FUNCTION_BLOCK STRING_TO_CAN_MSG (* STRING (bis 8 Zeichen) in eine CAN_MSG fuer AlPgnTxNew8B packen *)
  (* Standard: 61499-2; Description: Copyright (c) 2026 HR Agrartechnik GmbH This program and the accompanying materials are made available under the terms of the Eclipse Public License 2.0 which is available at https://www.eclipse.org/legal/epl-2.0/ SPDX-License-Identifier: EPL-2.0 *)
  (* Version 1.1, 2026-11-14, Franz Höpfinger, HR Agrartechnik GmbH, Fuellung Text + 16#00 + 16#FF, u16DaSize immer 8, PRIO auf 0..7 begrenzt, Ausgang TRUNC in TRUNCATED umbenannt (TRUNC ist reserviert) *)
  (* Version 1.0, 2026-11-13, Franz Höpfinger, HR Agrartechnik GmbH, Initial Version - STRING ueber CAN (0-8 Byte) *)
  PACKAGE isobus::pgn;
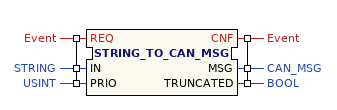
  EVENT_INPUT
    REQ WITH IN, PRIO; (* Text packen *)
  END_EVENT
  EVENT_OUTPUT
    CNF WITH MSG, TRUNCATED; (* MSG ist gefuellt *)
  END_EVENT
  VAR_INPUT
    IN : STRING; (* Text, je Zeichen 1 Byte *)
    PRIO : USINT := 6; (* Prioritaet (0..7), groesser 7 wird 7; AlPgnTxNew8B nimmt die Prioritaet vom install, nicht aus MSG *)
  END_VAR
  VAR_OUTPUT
    MSG : isobus::pgn::CAN_MSG; (* data = Zeichen, dann 16#00 (falls Platz), Rest 16#FF; u16DaSize = 8 *)
    TRUNCATED : BOOL; (* TRUE, wenn IN laenger als 8 Zeichen war (abgeschnitten) *)
  END_VAR
  EC_STATES
    REQ : REQ -> CNF;
  END_STATES
  ALGORITHM REQ IN ST: (* Zeichen in data[0..7] kopieren, mit 16#00 abschliessen, Rest 16#FF *)
VAR_TEMP
	n : DINT; // Anzahl zu kopierender Zeichen
	i : DINT; // Laufindex
END_VAR
n := LEN(IN);
IF n < 0 THEN
	n := 0;
END_IF;
TRUNCATED := n > 8;
IF n > 8 THEN
	n := 8;
END_IF;
FOR i := 0 TO 7 DO
	MSG.data[i] := BYTE#16#FF; // nicht genutzte Bytes wie bei J1939/ISOBUS ueblich
END_FOR;
FOR i := 1 TO n DO
	MSG.data[i - 1] := CHAR_TO_BYTE(IN[i]);
END_FOR;
IF n < 8 THEN
	MSG.data[n] := BYTE#16#00; // Textende
END_IF;
(* AlPgnTxNew8B sendet Laenge und Prioritaet vom install, MSG.u16DaSize und MSG.u8Priority werden dort nicht gelesen *)
MSG.u16DaSize := 8;
IF PRIO > 7 THEN
	MSG.u8Priority := 7;
ELSE
	MSG.u8Priority := PRIO;
END_IF;
  END_ALGORITHM
END_FUNCTION_BLOCK
